(* IEC 61131-3 sources: JingjiangMoonbox/Application/Application/数据类型/系统参数/站轴关系表, 2 files *)

(* ---- StAxisIdListInf.st ---- *)
(*@CES
Name=StAxisIdListInf
Type=Gvl
TypeGuid=2db5746d-d284-4425-9f7f-2663a34b0ebc
Guid=2e898926-372a-4322-a5eb-b0bb4f9f030f
HasDeclaration=True
HasImplementation=False
*)
{DECLARATION}
TYPE StAxisIdListInf :
STRUCT
	iAxisId: INT;(*轴号*)(*规划器*)
	iCoreId: int;(*核*)
	iTypeId: INT;(*类型*)
	iUnitId: INT;(*色组号*)
	iStdId: INT;(*站号*)
	iGroupId : INT;(*龙门组号*)
	iAdjAxisId : INT;(*调整轴号*)(*规划器*)
END_STRUCT
END_TYPE

{IMPLEMENTATION}

(* ---- StStationInfo_KS.st ---- *)
(*@CES
Name=StStationInfo_KS
Type=Gvl
TypeGuid=2db5746d-d284-4425-9f7f-2663a34b0ebc
Guid=6f2c3f0d-cedf-4320-89f1-935f04814eef
HasDeclaration=True
HasImplementation=False
*)
{DECLARATION}
TYPE StStationInfo_KS :
STRUCT
	iSid_Device: INT;
	iStationNum: INT;
	aiStationId_List: ARRAY [1..128] OF INT;(*设备站号*)
	awStation_Type: ARRAY [1..128] OF WORD;(*站类型*)
END_STRUCT
END_TYPE

{IMPLEMENTATION}
